(* IEC 61131-3 sources: model-first-plc-agent-ai/results/T2-W-19, 2 files *)

(* ---- a1_code.st ---- *)
FUNCTION_BLOCK FillingRuntime
VAR_INPUT
    start : BOOL;
    stop : BOOL;
    LSH : BOOL;
    LSHH : BOOL;
    TimerDuration : TIME;
END_VAR
VAR_OUTPUT
    fill_valve : BOOL;
    discharge_valve : BOOL;
END_VAR
VAR
    x0 : BOOL := TRUE;
    x1 : BOOL := FALSE;
    timer_done : BOOL := FALSE;
    FillingTimer : TON;
END_VAR

(* Evaluate the transition from the initial step. *)
IF x0 THEN
    IF start AND NOT stop AND NOT LSHH THEN
        x0 := FALSE;
        x1 := TRUE;
    END_IF;
END_IF;

(* Start timing in the scan in which the filling step becomes active. *)
FillingTimer(IN := x1, PT := TimerDuration);
timer_done := FillingTimer.Q;

(* Evaluate filling termination before assigning the physical outputs. *)
IF x1 THEN
    IF stop OR LSHH OR timer_done THEN
        x1 := FALSE;
        x0 := TRUE;

        (* Reset the step-owned timer immediately on leaving the step. *)
        FillingTimer(IN := FALSE, PT := TimerDuration);
        timer_done := FillingTimer.Q;
    END_IF;
END_IF;

fill_valve := x1;
discharge_valve := FALSE;

END_FUNCTION_BLOCK

PROGRAM Main
VAR
    StartCommand AT %IX100.0 : BOOL;
    StopCommand AT %IX100.1 : BOOL;
    LSH AT %IX100.2 : BOOL;
    LSHH AT %IX100.3 : BOOL;
    FillValve AT %QX100.0 : BOOL;
    DischargeValve AT %QX100.1 : BOOL;
END_VAR
VAR
    (* Configurable filling duration; adjust for the user scene. *)
    TimerDuration : TIME := T#10s;
    StartEdge : R_TRIG;
    RuntimeLogic : FillingRuntime;
END_VAR

StartEdge(CLK := StartCommand);

RuntimeLogic(
    start := StartEdge.Q,
    stop := StopCommand,
    LSH := LSH,
    LSHH := LSHH,
    TimerDuration := TimerDuration
);

FillValve := RuntimeLogic.fill_valve;
DischargeValve := RuntimeLogic.discharge_valve;

END_PROGRAM

(* ---- a2_code.st ---- *)
FUNCTION_BLOCK FB_TimedTankFilling
VAR_INPUT
    StartCommand : BOOL;
    StopCommand : BOOL;
    LSH : BOOL;
    LSHH : BOOL;
    TimerDuration : TIME;
END_VAR
VAR_OUTPUT
    fill_valve : BOOL;
    discharge_valve : BOOL;
END_VAR
VAR
    StartEdge : R_TRIG;
    FillingTimer : TON;
    SequenceState : INT := 0;
    start : BOOL;
    stop : BOOL;
    timer_done : BOOL;
END_VAR

StartEdge(CLK := StartCommand);
start := StartEdge.Q;
stop := StopCommand;

IF stop THEN
    SequenceState := 0;
ELSE
    CASE SequenceState OF
        0:
            IF start THEN
                SequenceState := 1;
            END_IF;
        1:
            SequenceState := 1;
    ELSE
        SequenceState := 0;
    END_CASE;
END_IF;

FillingTimer(
    IN := (SequenceState = 1),
    PT := TimerDuration
);
timer_done := FillingTimer.Q;

IF SequenceState = 1 THEN
    IF stop OR timer_done OR LSHH THEN
        SequenceState := 0;
    END_IF;
END_IF;

(* Reset the timer immediately on leaving the filling step. *)
IF SequenceState = 0 THEN
    FillingTimer(IN := FALSE, PT := TimerDuration);
    timer_done := FillingTimer.Q;
END_IF;

fill_valve := (SequenceState = 1) AND NOT stop;
discharge_valve := FALSE;

END_FUNCTION_BLOCK

PROGRAM Main
VAR
    StartCommand AT %IX100.0 : BOOL;
    StopCommand AT %IX100.1 : BOOL;
    LSH AT %IX100.2 : BOOL;
    LSHH AT %IX100.3 : BOOL;
    FillValve AT %QX100.0 : BOOL;
    DischargeValve AT %QX100.1 : BOOL;
END_VAR
VAR
    TankController : FB_TimedTankFilling;
    (* Configurable filling duration; adjust for the application. *)
    TimerDuration : TIME := T#5s;
END_VAR

TankController(
    StartCommand := StartCommand,
    StopCommand := StopCommand,
    LSH := LSH,
    LSHH := LSHH,
    TimerDuration := TimerDuration
);

FillValve := TankController.fill_valve;
DischargeValve := TankController.discharge_valve;

END_PROGRAM
